(*!
<summary>Selects one independently reported IO model test scenario.</summary>
*)
{attribute 'qualified_only'}
{attribute 'strict'}
TYPE IO_MODELS_TEST_SCENARIO :
(
	PULSE_TRAIN,
	ENCODER_CHANNELS,
	POWER_MEASUREMENT,
	AUXILIARY,
	COUNTER_AND_LOAD,
	SERIAL_AND_DIAGNOSTICS,
	DISCRETE_CATALOG,
	ANALOG_REPRESENTATIONS,
	DINT_BINDING,
	REAL_BINDING
);
END_TYPE

(* stored: Version 1.1.0.1
   DUT IO_MODELS_TEST_SCENARIO: Id {a51839d2-09e5-4fca-9ea4-822624370bf4} *)
